Fanuc KAREL source: KO00006.KL

PROGRAM KO00006
%NOLOCKGROUP
VAR
  P1: POSITION
  P2: POSITION
  P3: POSITION
  P4: POSITION
  OUT: XYZWPR
BEGIN
  OUT = FRAME(P1, P2, P3, P4)
END KO00006
